(* CODESYS project Overview.export

Project tree, tasks and I/O mapping:
  visualisation Overview
*)

// /Overview
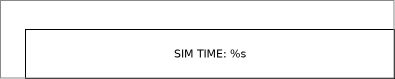
VISUALIZATION Overview  // 395x79
    Rectangle (25,29 370x50), "SIM TIME: %s", text variable: Team_HMI.sDateTime
END_VISUALIZATION
